Fanuc KAREL source: kd00072.KL

PROGRAM KD00072
%STACKSIZE=65535
%PRIORITY=65535
%NOLOCKGROUP
VAR
I : INTEGER
J : INTEGER
B : BOOLEAN
R : REAL
S : STRING[80]
BEGIN
-- UNRESOLVED_PC line 10 opcodes [9D 2E 1F] marker_code=0
END KD00072
